(* Tests FB_SpanProtoJsonSerializer: span fields, and grouping by resource and scope. *)
FUNCTION_BLOCK FB_TestSpanProtoJsonSerializer EXTENDS FB_TestSuite

THIS^.testSerializeRootSpan();
THIS^.testSerializeChildSpan();
THIS^.testSerializeSpanRejectsInvalidInput();
THIS^.testSerializeTracesDataWithEmptyQueue();
THIS^.testSerializeTracesDataGroupsByResourceAndScope();
THIS^.testSerializeSpanLinks();
THIS^.testSerializeLongTraceState();

(* A root span is written with hex identifiers, numeric enums, string timestamps, attributes and status, and no parentSpanId. *)
METHOD testSerializeRootSpan : REFERENCE TO FB_Test
VAR
	resource: FB_Resource('');
	idGenerator: FB_MockIdGenerator;
	provider: FB_TracerProvider_ForInspection(resource:=resource, idGenerator:=idGenerator, sampler:=TcOtlp_GVL.defaultSampler);
	scope: FB_InstrumentationScope('tracer.test', '1.0.0', '');
	tracer: FB_Tracer(scope:=scope, provider:=provider);
	serializer: FB_SpanProtoJsonSerializer;
	pSpan: POINTER TO FB_Span;
	root: SJsonValue;
	spans: SJsonValue;
	obj: SJsonValue;
	attribute: SJsonValue;
	status: SJsonValue;
	success: BOOL;
	reason: E_ProtoJsonSerializerFailureReason;
END_VAR
TcUnit.TEST('testSerializeRootSpan');
	tracer
		.startSpan(name:='work')
		.setStringAttribute(key:='stats.label', value:='pVal')
		.build(pDest:=pSpan);
	THIS^.AssertTrue(pSpan <> 0, 'Expected the span to build');
	IF pSpan <> 0 THEN
		// no builder sets timestamps; fixed values replace the clock so the output is known
		pSpan^.startTimestamp := 1000;
		pSpan^.endTimestamp := 1581452773000000789;
		tracer.setSpanStatusError(pSpan:=pSpan, message:='motor stalled');

		root := serializer.parser.NewDocument();
		root := serializer.parser.SetObject(root);
		spans := serializer.parser.AddArrayMember(root, 'spans', 0);
		success := serializer.serializeSpan(v:=spans, pSpan:=pSpan, failureReason=>reason);
		THIS^.AssertTrue(success, 'Expected the span to serialize');
		THIS^.AssertEquals_UDINT(TO_UDINT(E_ProtoJsonSerializerFailureReason.NA), TO_UDINT(reason), 'Expected no failure reason');

		obj := serializer.parser.GetArrayValueByIdx(spans, 0);
		THIS^.AssertTrue(serializer.parser.IsObject(obj), 'Expected one Span object');
		// FB_MockIdGenerator fills each new id with one counter byte: the trace id gets 01, the span id 02
		THIS^.AssertEquals_STRING('01010101010101010101010101010101', serializer.parser.GetString(serializer.parser.FindMember(obj, 'traceId')), 'Expected the hex traceId');
		THIS^.AssertEquals_STRING('0202020202020202', serializer.parser.GetString(serializer.parser.FindMember(obj, 'spanId')), 'Expected the hex spanId');
		THIS^.AssertTrue(serializer.parser.FindMember(obj, 'parentSpanId') = 0, 'Expected a root span to omit parentSpanId');
		THIS^.AssertEquals_STRING('work', serializer.parser.GetString(serializer.parser.FindMember(obj, 'name')), 'Expected the name');
		THIS^.AssertEquals_UDINT(1, serializer.parser.GetUint(serializer.parser.FindMember(obj, 'kind')), 'Expected SPAN_KIND_INTERNAL as a number');
		THIS^.AssertEquals_STRING('1000', serializer.parser.GetString(serializer.parser.FindMember(obj, 'startTimeUnixNano')), 'Expected a string startTimeUnixNano');
		THIS^.AssertEquals_STRING('1581452773000000789', serializer.parser.GetString(serializer.parser.FindMember(obj, 'endTimeUnixNano')), 'Expected a string endTimeUnixNano');

		attribute := serializer.parser.GetArrayValueByIdx(serializer.parser.FindMember(obj, 'attributes'), 0);
		THIS^.AssertEquals_STRING('stats.label', serializer.parser.GetString(serializer.parser.FindMember(attribute, 'key')), 'Expected the attribute key');
		THIS^.AssertEquals_STRING(
			'pVal',
			serializer.parser.GetString(serializer.parser.FindMember(serializer.parser.FindMember(attribute, 'value'), 'stringValue')),
			'Expected the attribute value'
		);

		status := serializer.parser.FindMember(obj, 'status');
		THIS^.AssertEquals_UDINT(2, serializer.parser.GetUint(serializer.parser.FindMember(status, 'code')), 'Expected STATUS_CODE_ERROR as a number');
		THIS^.AssertEquals_STRING('motor stalled', serializer.parser.GetString(serializer.parser.FindMember(status, 'message')), 'Expected the status message');
		THIS^.AssertTrue(pSpan^.name <> 0 AND_THEN pSpan^.status <> 0, 'Expected serialization to leave the span intact');
	END_IF

	IF pSpan <> 0 THEN pSpan^.delete(pSelf:=pSpan); END_IF
TcUnit.TEST_FINISHED();
END_METHOD

(* A child span is written with its parentSpanId and kind, and without a status when none is set. *)
METHOD testSerializeChildSpan : REFERENCE TO FB_Test
VAR
	resource: FB_Resource('');
	idGenerator: FB_MockIdGenerator;
	provider: FB_TracerProvider_ForInspection(resource:=resource, idGenerator:=idGenerator, sampler:=TcOtlp_GVL.defaultSampler);
	scope: FB_InstrumentationScope('tracer.test', '1.0.0', '');
	tracer: FB_Tracer(scope:=scope, provider:=provider);
	serializer: FB_SpanProtoJsonSerializer;
	pRoot: POINTER TO FB_Span;
	pChild: POINTER TO FB_Span;
	pContext: POINTER TO FB_SpanContext;
	root: SJsonValue;
	spans: SJsonValue;
	obj: SJsonValue;
	success: BOOL;
END_VAR
TcUnit.TEST('testSerializeChildSpan');
	tracer.startSpan(name:='root').build(pDest:=pRoot);
	IF pRoot <> 0 THEN
		tracer.getSpanContext(pSpan:=pRoot, pDest:=pContext);
	END_IF
	tracer
		.startSpan(name:='child', kind:=E_SpanKind.SPAN_KIND_CLIENT)
		.setParentUsingContext(pContext:=pContext)
		.build(pDest:=pChild);
	THIS^.AssertTrue(pChild <> 0, 'Expected the child span to build');
	IF pChild <> 0 THEN
		root := serializer.parser.NewDocument();
		root := serializer.parser.SetObject(root);
		spans := serializer.parser.AddArrayMember(root, 'spans', 0);
		success := serializer.serializeSpan(v:=spans, pSpan:=pChild);
		THIS^.AssertTrue(success, 'Expected the child span to serialize');

		obj := serializer.parser.GetArrayValueByIdx(spans, 0);
		// FB_MockIdGenerator fills each new id with one counter byte: the root takes trace 01 and
		// span 02, and the child keeps the root's trace and takes span 03
		THIS^.AssertEquals_STRING('0303030303030303', serializer.parser.GetString(serializer.parser.FindMember(obj, 'spanId')), 'Expected the child spanId');
		THIS^.AssertEquals_STRING('0202020202020202', serializer.parser.GetString(serializer.parser.FindMember(obj, 'parentSpanId')), 'Expected the parent spanId');
		THIS^.AssertEquals_UDINT(3, serializer.parser.GetUint(serializer.parser.FindMember(obj, 'kind')), 'Expected SPAN_KIND_CLIENT as a number');
		THIS^.AssertTrue(serializer.parser.FindMember(obj, 'status') = 0, 'Expected no status member');
		THIS^.AssertTrue(serializer.parser.FindMember(obj, 'attributes') = 0, 'Expected no attributes member');
	END_IF

	IF pContext <> 0 THEN pContext^.delete(pSelf:=pContext); END_IF
	IF pChild <> 0 THEN pChild^.delete(pSelf:=pChild); END_IF
	IF pRoot <> 0 THEN pRoot^.delete(pSelf:=pRoot); END_IF
TcUnit.TEST_FINISHED();
END_METHOD

(* serializeSpan reports a null span and an invalid JSON destination. *)
METHOD testSerializeSpanRejectsInvalidInput : REFERENCE TO FB_Test
VAR
	resource: FB_Resource('');
	idGenerator: FB_MockIdGenerator;
	provider: FB_TracerProvider_ForInspection(resource:=resource, idGenerator:=idGenerator, sampler:=TcOtlp_GVL.defaultSampler);
	scope: FB_InstrumentationScope('tracer.test', '1.0.0', '');
	tracer: FB_Tracer(scope:=scope, provider:=provider);
	serializer: FB_SpanProtoJsonSerializer;
	root: SJsonValue;
	spans: SJsonValue;
	invalid: SJsonValue;
	pSpan: POINTER TO FB_Span;
	success: BOOL;
	reason: E_ProtoJsonSerializerFailureReason;
END_VAR
TcUnit.TEST('testSerializeSpanRejectsInvalidInput');
	root := serializer.parser.NewDocument();
	root := serializer.parser.SetObject(root);
	spans := serializer.parser.AddArrayMember(root, 'spans', 0);

	success := serializer.serializeSpan(v:=spans, pSpan:=pSpan, failureReason=>reason);
	THIS^.AssertFalse(success, 'Expected a null span to fail');
	THIS^.AssertEquals_UDINT(TO_UDINT(E_ProtoJsonSerializerFailureReason.SPAN_POINTER_NULL), TO_UDINT(reason), 'Expected SPAN_POINTER_NULL');

	// a valid span, so the only fault left is the destination, which invalid leaves at 0
	tracer.startSpan(name:='work').build(pDest:=pSpan);
	THIS^.AssertTrue(pSpan <> 0, 'Expected the span to build');
	success := serializer.serializeSpan(v:=invalid, pSpan:=pSpan, failureReason=>reason);
	THIS^.AssertFalse(success, 'Expected an invalid destination to fail');
	THIS^.AssertEquals_UDINT(TO_UDINT(E_ProtoJsonSerializerFailureReason.JSON_VALUE_INVALID), TO_UDINT(reason), 'Expected JSON_VALUE_INVALID');
	IF pSpan <> 0 THEN pSpan^.delete(pSelf:=pSpan); END_IF
TcUnit.TEST_FINISHED();
END_METHOD

(* An empty queue gives a document with an empty resourceSpans array. *)
METHOD testSerializeTracesDataWithEmptyQueue : REFERENCE TO FB_Test
VAR
	serializer: FB_SpanProtoJsonSerializer;
	queue: FB_SpanQueue(maxCount:=0);
	resourceSpans: SJsonValue;
	success: BOOL;
	reason: E_ProtoJsonSerializerFailureReason;
END_VAR
TcUnit.TEST('testSerializeTracesDataWithEmptyQueue');
	success := serializer.serializeTracesData(spans:=queue, failureReason=>reason);
	THIS^.AssertTrue(success, 'Expected an empty queue to serialize');
	THIS^.AssertEquals_UDINT(TO_UDINT(E_ProtoJsonSerializerFailureReason.NA), TO_UDINT(reason), 'Expected no failure reason');
	resourceSpans := serializer.parser.FindMember(serializer.jsonValue, 'resourceSpans');
	THIS^.AssertTrue(resourceSpans <> 0 AND_THEN serializer.parser.IsArray(resourceSpans), 'Expected a resourceSpans array');
	THIS^.AssertTrue(serializer.parser.GetArrayValueByIdx(resourceSpans, 0) = 0, 'Expected no ResourceSpans groups');
TcUnit.TEST_FINISHED();
END_METHOD

(*
	Spans arrive with interleaved resources and scopes. Each resource is written once with
	its scopes in first-seen order, and spans keep queue order inside a scope. The serializer
	drains the queue, releasing every span.
*)
METHOD testSerializeTracesDataGroupsByResourceAndScope : REFERENCE TO FB_Test
VAR
	idGenerator: FB_MockIdGenerator;
	resourceB: FB_Resource('resource.b');
	resourceA: FB_Resource('resource.a');
	resourceC: FB_Resource('resource.c');
	providerB: FB_TracerProvider_ForInspection(resource:=resourceB, idGenerator:=idGenerator, sampler:=TcOtlp_GVL.defaultSampler);
	providerA: FB_TracerProvider_ForInspection(resource:=resourceA, idGenerator:=idGenerator, sampler:=TcOtlp_GVL.defaultSampler);
	providerC: FB_TracerProvider_ForInspection(resource:=resourceC, idGenerator:=idGenerator, sampler:=TcOtlp_GVL.defaultSampler);
	scopeB: FB_InstrumentationScope('scope.b', '1.0.0', 'scope.b.schema');
	scopeA: FB_InstrumentationScope('scope.a', '1.0.0', 'scope.a.schema');
	scopeC: FB_InstrumentationScope('scope.c', '1.0.0', 'scope.c.schema');
	tracerBb: FB_Tracer(scope:=scopeB, provider:=providerB);
	tracerBa: FB_Tracer(scope:=scopeA, provider:=providerB);
	tracerAc: FB_Tracer(scope:=scopeC, provider:=providerA);
	tracerAb: FB_Tracer(scope:=scopeB, provider:=providerA);
	tracerCa: FB_Tracer(scope:=scopeA, provider:=providerC);
	queue: FB_SpanQueue(maxCount:=0);
	serializer: FB_SpanProtoJsonSerializer;
	pSpan: POINTER TO FB_Span;
	name: T_MaxString;
	idx: UDINT;
	success: BOOL;
	reason: E_ProtoJsonSerializerFailureReason;
	resourceSpans: SJsonValue;
	resourceObj: SJsonValue;
	scopeSpans: SJsonValue;
	scopeObj: SJsonValue;
	spanArray: SJsonValue;
	spanObj: SJsonValue;
END_VAR
TcUnit.TEST('testSerializeTracesDataGroupsByResourceAndScope');
	// ---- Arrange: eight spans with interleaved resource/scope pairs ----
	// Each tracer is one resource/scope pair, named resource then scope (tracerBa is resource B, scope A).
	// The name holds the span number, so each span can be identified in the output.
	//   span:     1  2  3  4  5  6  7  8
	//   resource: B  A  C  B  C  A  B  A
	//   scope:    B  C  A  A  A  B  B  C
	FOR idx := 1 TO 8 DO
		name := CONCAT('span', UDINT_TO_STRING(idx));
		CASE idx OF
			1, 7: tracerBb.startSpan(name:=name).build(pDest:=pSpan);
			4: tracerBa.startSpan(name:=name).build(pDest:=pSpan);
			2, 8: tracerAc.startSpan(name:=name).build(pDest:=pSpan);
			6: tracerAb.startSpan(name:=name).build(pDest:=pSpan);
			3, 5: tracerCa.startSpan(name:=name).build(pDest:=pSpan);
		END_CASE
		THIS^.AssertTrue(pSpan <> 0, CONCAT('Expected to build ', name));
		IF pSpan <> 0 AND_THEN NOT queue.push(pValue:=pSpan) THEN
			pSpan^.delete(pSelf:=pSpan);
		END_IF
	END_FOR
	THIS^.AssertEquals_UDINT(8, queue.count, 'Expected eight queued spans');

	// ---- Act ----
	success := serializer.serializeTracesData(spans:=queue, failureReason=>reason);
	THIS^.AssertTrue(success, 'Expected TracesData to serialize');
	THIS^.AssertEquals_UDINT(TO_UDINT(E_ProtoJsonSerializerFailureReason.NA), TO_UDINT(reason), 'Expected no failure reason');
	THIS^.AssertEquals_UDINT(0, queue.count, 'Expected the serializer to drain the queue');
	resourceSpans := serializer.parser.FindMember(serializer.jsonValue, 'resourceSpans');
	THIS^.AssertTrue(resourceSpans <> 0 AND_THEN serializer.parser.IsArray(resourceSpans), 'Expected a resourceSpans array');
	THIS^.AssertTrue(serializer.parser.GetArrayValueByIdx(resourceSpans, 3) = 0, 'Expected exactly three ResourceSpans groups');

	// ---- Assert: resource B was seen first, with scope B (spans 1, 7) before scope A (span 4) ----
	resourceObj := serializer.parser.GetArrayValueByIdx(resourceSpans, 0);
	THIS^.AssertEquals_STRING('resource.b', serializer.parser.GetString(serializer.parser.FindMember(resourceObj, 'schemaUrl')), 'Expected resource.b at 0');
	scopeSpans := serializer.parser.FindMember(resourceObj, 'scopeSpans');
	scopeObj := serializer.parser.GetArrayValueByIdx(scopeSpans, 0);
	THIS^.AssertEquals_STRING('scope.b', serializer.parser.GetString(serializer.parser.FindMember(serializer.parser.FindMember(scopeObj, 'scope'), 'name')), 'Expected resource.b scope.b at 0');
	spanArray := serializer.parser.FindMember(scopeObj, 'spans');
	spanObj := serializer.parser.GetArrayValueByIdx(spanArray, 0);
	THIS^.AssertEquals_STRING('span1', serializer.parser.GetString(serializer.parser.FindMember(spanObj, 'name')), 'Expected span1 in resource.b scope.b');
	spanObj := serializer.parser.GetArrayValueByIdx(spanArray, 1);
	THIS^.AssertEquals_STRING('span7', serializer.parser.GetString(serializer.parser.FindMember(spanObj, 'name')), 'Expected span7 in resource.b scope.b');
	THIS^.AssertTrue(serializer.parser.GetArrayValueByIdx(spanArray, 2) = 0, 'Expected 2 span(s) in resource.b scope.b');

	scopeObj := serializer.parser.GetArrayValueByIdx(scopeSpans, 1);
	THIS^.AssertEquals_STRING('scope.a', serializer.parser.GetString(serializer.parser.FindMember(serializer.parser.FindMember(scopeObj, 'scope'), 'name')), 'Expected resource.b scope.a at 1');
	spanArray := serializer.parser.FindMember(scopeObj, 'spans');
	spanObj := serializer.parser.GetArrayValueByIdx(spanArray, 0);
	THIS^.AssertEquals_STRING('span4', serializer.parser.GetString(serializer.parser.FindMember(spanObj, 'name')), 'Expected span4 in resource.b scope.a');
	THIS^.AssertTrue(serializer.parser.GetArrayValueByIdx(spanArray, 1) = 0, 'Expected 1 span(s) in resource.b scope.a');
	THIS^.AssertTrue(serializer.parser.GetArrayValueByIdx(scopeSpans, 2) = 0, 'Expected 2 scope(s) in resource.b');

	// resource A was seen second, with scope C (spans 2, 8) before scope B (span 6)
	resourceObj := serializer.parser.GetArrayValueByIdx(resourceSpans, 1);
	THIS^.AssertEquals_STRING('resource.a', serializer.parser.GetString(serializer.parser.FindMember(resourceObj, 'schemaUrl')), 'Expected resource.a at 1');
	scopeSpans := serializer.parser.FindMember(resourceObj, 'scopeSpans');
	scopeObj := serializer.parser.GetArrayValueByIdx(scopeSpans, 0);
	THIS^.AssertEquals_STRING('scope.c', serializer.parser.GetString(serializer.parser.FindMember(serializer.parser.FindMember(scopeObj, 'scope'), 'name')), 'Expected resource.a scope.c at 0');
	spanArray := serializer.parser.FindMember(scopeObj, 'spans');
	spanObj := serializer.parser.GetArrayValueByIdx(spanArray, 0);
	THIS^.AssertEquals_STRING('span2', serializer.parser.GetString(serializer.parser.FindMember(spanObj, 'name')), 'Expected span2 in resource.a scope.c');
	spanObj := serializer.parser.GetArrayValueByIdx(spanArray, 1);
	THIS^.AssertEquals_STRING('span8', serializer.parser.GetString(serializer.parser.FindMember(spanObj, 'name')), 'Expected span8 in resource.a scope.c');
	THIS^.AssertTrue(serializer.parser.GetArrayValueByIdx(spanArray, 2) = 0, 'Expected 2 span(s) in resource.a scope.c');

	scopeObj := serializer.parser.GetArrayValueByIdx(scopeSpans, 1);
	THIS^.AssertEquals_STRING('scope.b', serializer.parser.GetString(serializer.parser.FindMember(serializer.parser.FindMember(scopeObj, 'scope'), 'name')), 'Expected resource.a scope.b at 1');
	spanArray := serializer.parser.FindMember(scopeObj, 'spans');
	spanObj := serializer.parser.GetArrayValueByIdx(spanArray, 0);
	THIS^.AssertEquals_STRING('span6', serializer.parser.GetString(serializer.parser.FindMember(spanObj, 'name')), 'Expected span6 in resource.a scope.b');
	THIS^.AssertTrue(serializer.parser.GetArrayValueByIdx(spanArray, 1) = 0, 'Expected 1 span(s) in resource.a scope.b');
	THIS^.AssertTrue(serializer.parser.GetArrayValueByIdx(scopeSpans, 2) = 0, 'Expected 2 scope(s) in resource.a');

	// resource C was seen third; its non-adjacent spans 3 and 5 share scope A
	resourceObj := serializer.parser.GetArrayValueByIdx(resourceSpans, 2);
	THIS^.AssertEquals_STRING('resource.c', serializer.parser.GetString(serializer.parser.FindMember(resourceObj, 'schemaUrl')), 'Expected resource.c at 2');
	scopeSpans := serializer.parser.FindMember(resourceObj, 'scopeSpans');
	scopeObj := serializer.parser.GetArrayValueByIdx(scopeSpans, 0);
	THIS^.AssertEquals_STRING('scope.a', serializer.parser.GetString(serializer.parser.FindMember(serializer.parser.FindMember(scopeObj, 'scope'), 'name')), 'Expected resource.c scope.a at 0');
	spanArray := serializer.parser.FindMember(scopeObj, 'spans');
	spanObj := serializer.parser.GetArrayValueByIdx(spanArray, 0);
	THIS^.AssertEquals_STRING('span3', serializer.parser.GetString(serializer.parser.FindMember(spanObj, 'name')), 'Expected span3 in resource.c scope.a');
	spanObj := serializer.parser.GetArrayValueByIdx(spanArray, 1);
	THIS^.AssertEquals_STRING('span5', serializer.parser.GetString(serializer.parser.FindMember(spanObj, 'name')), 'Expected span5 in resource.c scope.a');
	THIS^.AssertTrue(serializer.parser.GetArrayValueByIdx(spanArray, 2) = 0, 'Expected 2 span(s) in resource.c scope.a');
	THIS^.AssertTrue(serializer.parser.GetArrayValueByIdx(scopeSpans, 1) = 0, 'Expected 1 scope(s) in resource.c');

	queue.free();
TcUnit.TEST_FINISHED();
END_METHOD

(* Links are written as a 'links' array in the order they were added, each with hex
   identifiers, flags and any attributes. A span without links writes no 'links' member. *)
METHOD testSerializeSpanLinks : REFERENCE TO FB_Test
VAR
	resource: FB_Resource('');
	idGenerator: FB_MockIdGenerator;
	provider: FB_TracerProvider_ForInspection(resource:=resource, idGenerator:=idGenerator, sampler:=TcOtlp_GVL.defaultSampler);
	scope: FB_InstrumentationScope('tracer.test', '1.0.0', '');
	tracer: FB_Tracer(scope:=scope, provider:=provider);
	serializer: FB_SpanProtoJsonSerializer;
	pTrigger: POINTER TO FB_Span;
	pSpan: POINTER TO FB_Span;
	pTriggerContext: POINTER TO FB_SpanContext;
	pLink: POINTER TO FB_Link;
	root: SJsonValue;
	spans: SJsonValue;
	obj: SJsonValue;
	links: SJsonValue;
	link: SJsonValue;
	attribute: SJsonValue;
	success: BOOL;
	reason: E_ProtoJsonSerializerFailureReason;
END_VAR
TcUnit.TEST('testSerializeSpanLinks');
	tracer.startSpan(name:='trigger').build(pDest:=pTrigger);
	IF pTrigger <> 0 THEN tracer.getSpanContext(pSpan:=pTrigger, pDest:=pTriggerContext); END_IF
	tracer.startSpan(name:='work').addLink(pContext:=pTriggerContext).build(pDest:=pSpan);
	THIS^.AssertTrue(pSpan <> 0, 'Expected the linked span to build');

	// a link with attributes is built with LinkFactory and pushed to the running span
	LinkFactory.fromSpan(pDest:=pLink, pSpan:=pTrigger);
	IF pLink <> 0 THEN
		pLink^.attributes.setStringAttribute(key:='link.reason', value:='retry');
	END_IF
	tracer.pushSpanLink(pSpan:=pSpan, pLink:=pLink);

	IF pSpan <> 0 AND pTrigger <> 0 THEN
		root := serializer.parser.NewDocument();
		root := serializer.parser.SetObject(root);
		spans := serializer.parser.AddArrayMember(root, 'spans', 0);
		success := serializer.serializeSpan(v:=spans, pSpan:=pSpan, failureReason=>reason);
		THIS^.AssertTrue(success, 'Expected the linked span to serialize');
		THIS^.AssertEquals_UDINT(TO_UDINT(E_ProtoJsonSerializerFailureReason.NA), TO_UDINT(reason), 'Expected no failure reason');
		success := serializer.serializeSpan(v:=spans, pSpan:=pTrigger, failureReason=>reason);
		THIS^.AssertTrue(success, 'Expected the trigger span to serialize');

		obj := serializer.parser.GetArrayValueByIdx(spans, 0);
		links := serializer.parser.FindMember(obj, 'links');
		THIS^.AssertTrue(serializer.parser.IsArray(links), 'Expected a links array');
		THIS^.AssertTrue(serializer.parser.FindMember(obj, 'droppedLinksCount') = 0, 'Expected no droppedLinksCount when nothing was dropped');

		link := serializer.parser.GetArrayValueByIdx(links, 0);
		THIS^.AssertTrue(serializer.parser.IsObject(link), 'Expected the first Link object');
		// FB_MockIdGenerator fills each new id with one counter byte: the trigger took trace 01 and span 02
		THIS^.AssertEquals_STRING('01010101010101010101010101010101', serializer.parser.GetString(serializer.parser.FindMember(link, 'traceId')), 'Expected the hex linked traceId');
		THIS^.AssertEquals_STRING('0202020202020202', serializer.parser.GetString(serializer.parser.FindMember(link, 'spanId')), 'Expected the hex linked spanId');
		THIS^.AssertEquals_UDINT(16#101, serializer.parser.GetUint(serializer.parser.FindMember(link, 'flags')), 'Expected the sampled bit and a known local context (16#101)');
		THIS^.AssertTrue(serializer.parser.FindMember(link, 'attributes') = 0, 'Expected no attributes on the first link');
		THIS^.AssertTrue(serializer.parser.FindMember(link, 'traceState') = 0, 'Expected no traceState on the first link');

		link := serializer.parser.GetArrayValueByIdx(links, 1);
		THIS^.AssertTrue(serializer.parser.IsObject(link), 'Expected the second Link object');
		attribute := serializer.parser.GetArrayValueByIdx(serializer.parser.FindMember(link, 'attributes'), 0);
		THIS^.AssertEquals_STRING('link.reason', serializer.parser.GetString(serializer.parser.FindMember(attribute, 'key')), 'Expected the link attribute key');
		THIS^.AssertEquals_STRING(
			'retry',
			serializer.parser.GetString(serializer.parser.FindMember(serializer.parser.FindMember(attribute, 'value'), 'stringValue')),
			'Expected the link attribute value'
		);

		obj := serializer.parser.GetArrayValueByIdx(spans, 1);
		THIS^.AssertTrue(serializer.parser.FindMember(obj, 'links') = 0, 'Expected a span without links to omit links');
	END_IF

	IF pLink <> 0 THEN pLink^.delete(pSelf:=pLink); END_IF
	IF pTriggerContext <> 0 THEN pTriggerContext^.delete(pSelf:=pTriggerContext); END_IF
	IF pSpan <> 0 THEN pSpan^.delete(pSelf:=pSpan); END_IF
	IF pTrigger <> 0 THEN pTrigger^.delete(pSelf:=pTrigger); END_IF
TcUnit.TEST_FINISHED();
END_METHOD

(* A trace state longer than T_MaxString is written whole. W3C asks for at least 512 characters. *)
METHOD testSerializeLongTraceState : REFERENCE TO FB_Test
VAR
	resource: FB_Resource('');
	idGenerator: FB_MockIdGenerator;
	provider: FB_TracerProvider_ForInspection(resource:=resource, idGenerator:=idGenerator, sampler:=TcOtlp_GVL.defaultSampler);
	scope: FB_InstrumentationScope('tracer.test', '1.0.0', '');
	tracer: FB_Tracer(scope:=scope, provider:=provider);
	serializer: FB_SpanProtoJsonSerializer;
	header: STRING(600);
	written: STRING(600);
	pWritten: POINTER TO STRING;
	pBytes: POINTER TO BYTE;
	entry: UDINT;
	i: UDINT;
	n: UDINT;
	traceId: FB_TraceId;
	spanId: FB_SpanId;
	pTraceState: POINTER TO FB_TraceState;
	pRemote: POINTER TO FB_SpanContext;
	pSpan: POINTER TO FB_Span;
	root: SJsonValue;
	spans: SJsonValue;
	obj: SJsonValue;
	member: SJsonValue;
	success: BOOL;
	reason: E_ProtoJsonSerializerFailureReason;
END_VAR
TcUnit.TEST('testSerializeLongTraceState');
	// four 128 character entries joined by ',': 515 characters, built byte by byte
	pBytes := ADR(header);
	FOR entry := 0 TO 3 DO
		IF entry > 0 THEN
			pBytes[n] := 16#2C;  // ','
			n := n + 1;
		END_IF
		pBytes[n] := 16#6B;  // 'k'
		pBytes[n + 1] := 16#30 + TO_BYTE(entry);  // '0' to '3'
		pBytes[n + 2] := 16#3D;  // '='
		n := n + 3;
		FOR i := 1 TO 125 DO  // 125 value characters make a 128 character entry
			pBytes[n] := 16#61 + TO_BYTE(i MOD 26);  // 'a' to 'z'
			n := n + 1;
		END_FOR
	END_FOR
	pBytes[n] := 0;

	MEMSET(ADR(traceId.bytes), 16#AA, SIZEOF(traceId.bytes));
	MEMSET(ADR(spanId.bytes), 16#BB, SIZEOF(spanId.bytes));
	TraceStateFactory.parse(pDest:=pTraceState, pHeader:=ADR(header));
	// 16#301: sampled, remoteness known, remote
	ContextFactory.buildContext(pDest:=pRemote, pTraceId:=ADR(traceId), pSpanId:=ADR(spanId), pTraceState:=pTraceState, traceFlags:=16#301);
	IF pTraceState <> 0 THEN pTraceState^.delete(pSelf:=pTraceState); END_IF
	tracer.startSpan(name:='remote.child').setParentUsingContext(pContext:=pRemote).build(pDest:=pSpan);
	IF pRemote <> 0 THEN pRemote^.delete(pSelf:=pRemote); END_IF
	THIS^.AssertTrue(pSpan <> 0, 'Expected the span to build');

	IF pSpan <> 0 THEN
		root := serializer.parser.NewDocument();
		root := serializer.parser.SetObject(root);
		spans := serializer.parser.AddArrayMember(root, 'spans', 0);
		success := serializer.serializeSpan(v:=spans, pSpan:=pSpan, failureReason=>reason);
		THIS^.AssertTrue(success, 'Expected the span to serialize');

		obj := serializer.parser.GetArrayValueByIdx(spans, 0);
		member := serializer.parser.FindMember(obj, 'traceState');
		THIS^.AssertTrue(member <> 0, 'Expected a traceState member');
		IF member <> 0 THEN
			THIS^.AssertEquals_UDINT(516, TO_UDINT(serializer.parser.GetStringLength(member)), 'Expected all 515 characters and the terminator');
			pWritten := ADR(written);  // CopyString takes a STRING reference and a size, so it can fill a longer buffer
			serializer.parser.CopyString(member, pWritten^, SIZEOF(written));
			THIS^.AssertTrue(MEMCMP(ADR(written), ADR(header), 516) = 0, 'Expected the trace state unchanged');
		END_IF
		pSpan^.delete(pSelf:=pSpan);
	END_IF
TcUnit.TEST_FINISHED();
END_METHOD

END_FUNCTION_BLOCK

(* stored: Version 1.1.0.1
   POU FB_TestSpanProtoJsonSerializer: Id {db065884-1d07-4f0b-9eec-d553d5215051}, SpecialFunc None
   Method testSerializeRootSpan: Id {ffa2cc14-29c0-48dc-aa0d-c692404b304a}
   Method testSerializeChildSpan: Id {59235f6e-3375-4031-9daa-7f676956041d}
   Method testSerializeSpanRejectsInvalidInput: Id {12720abc-a60a-4ca1-9f13-38711b9d2830}
   Method testSerializeTracesDataWithEmptyQueue: Id {ca74d4ca-6f40-4128-b7c0-a7cc66b4ec06}
   Method testSerializeTracesDataGroupsByResourceAndScope: Id {9bcd3ce8-bfe8-48e7-ab1d-e1f108e0e7a3}
   Method testSerializeSpanLinks: Id {a9a9dda3-91e8-40bf-b4e7-2147740c442f}
   Method testSerializeLongTraceState: Id {fbe0bb89-4af4-4c50-8460-2f8ec01cc66c} *)
